Fanuc KAREL source: KA00023.KL

PROGRAM KA00023
%NOLOCKGROUP
VAR
  SRC: REAL
  DST: ARRAY[2] OF BYTE
BEGIN
  SRC = 2.0
  DST[1] = SRC
END KA00023
